(* IEC 61131-3 sources: plcassist-cli/packages/volt-lsp-iec/test-corpus/CodesysTestProject/Device/Plc Logic/Application/Library Manager/Standard, 22 files *)

(* ---- CONCAT.fun ---- *)
FUNCTION CONCAT : STRING(255)
VAR_INPUT
	STR1 : STRING(255);
	STR2 : STRING(255);
END_VAR
END_FUNCTION

(* ---- DELETE.fun ---- *)
FUNCTION DELETE : STRING(255)
VAR_INPUT
	STR : STRING(255);
	LEN : INT;
	POS : INT;
END_VAR
END_FUNCTION

(* ---- FIND.fun ---- *)
FUNCTION FIND : INT
VAR_INPUT
	STR1 : STRING(255);
	STR2 : STRING(255);
END_VAR
END_FUNCTION

(* ---- INSERT.fun ---- *)
FUNCTION INSERT : STRING(255)
VAR_INPUT
	STR1 : STRING(255);
	STR2 : STRING(255);
	POS : INT;
END_VAR
END_FUNCTION

(* ---- LEFT.fun ---- *)
FUNCTION LEFT : STRING(255)
VAR_INPUT
	STR : STRING(255);
	SIZE : INT;
END_VAR
END_FUNCTION

(* ---- LEN.fun ---- *)
FUNCTION LEN : INT
VAR_INPUT
	STR : STRING(255);
END_VAR
END_FUNCTION

(* ---- LEN_INTERNAL.fun ---- *)
FUNCTION LEN_INTERNAL : UINT
VAR_IN_OUT
	STR : STRING(255);
END_VAR
END_FUNCTION

(* ---- MEMCOPY_INTERNAL.fun ---- *)
FUNCTION MEMCOPY_INTERNAL : POINTER TO BYTE
VAR_INPUT
	PDEST : POINTER TO BYTE;
	PSRC : POINTER TO BYTE;
	DWSIZE : DWORD;
END_VAR
END_FUNCTION

(* ---- MID.fun ---- *)
FUNCTION MID : STRING(255)
VAR_INPUT
	STR : STRING(255);
	LEN : INT;
	POS : INT;
END_VAR
END_FUNCTION

(* ---- REPLACE.fun ---- *)
FUNCTION REPLACE : STRING(255)
VAR_INPUT
	STR1 : STRING(255);
	STR2 : STRING(255);
	L : INT;
	P : INT;
END_VAR
END_FUNCTION

(* ---- RIGHT.fun ---- *)
FUNCTION RIGHT : STRING(255)
VAR_INPUT
	STR : STRING(255);
	SIZE : INT;
END_VAR
END_FUNCTION

(* ---- CTD.fb ---- *)
FUNCTION_BLOCK CTD
VAR_INPUT
	CD : BOOL;
	LOAD : BOOL;
	PV : WORD;
END_VAR
VAR_OUTPUT
	Q : BOOL;
	CV : WORD;
END_VAR
VAR
	M : BOOL;
END_VAR
END_FUNCTION_BLOCK

(* ---- CTU.fb ---- *)
FUNCTION_BLOCK CTU
VAR_INPUT
	CU : BOOL;
	RESET : BOOL;
	PV : WORD;
END_VAR
VAR_OUTPUT
	Q : BOOL;
	CV : WORD;
END_VAR
VAR
	M : BOOL;
END_VAR
END_FUNCTION_BLOCK

(* ---- CTUD.fb ---- *)
FUNCTION_BLOCK CTUD
VAR_INPUT
	CU : BOOL;
	CD : BOOL;
	RESET : BOOL;
	LOAD : BOOL;
	PV : WORD;
END_VAR
VAR_OUTPUT
	QU : BOOL;
	QD : BOOL;
	CV : WORD;
END_VAR
VAR
	MU : BOOL;
	MD : BOOL;
	RU : BOOL;
	RD : BOOL;
END_VAR
END_FUNCTION_BLOCK

(* ---- F_TRIG.fb ---- *)
FUNCTION_BLOCK F_TRIG
VAR_INPUT
	CLK : BOOL;
END_VAR
VAR_OUTPUT
	Q : BOOL;
END_VAR
VAR
	M : BOOL := TRUE;
END_VAR
END_FUNCTION_BLOCK

(* ---- R_TRIG.fb ---- *)
FUNCTION_BLOCK R_TRIG
VAR_INPUT
	CLK : BOOL;
END_VAR
VAR_OUTPUT
	Q : BOOL;
END_VAR
VAR
	M : BOOL;
END_VAR
END_FUNCTION_BLOCK

(* ---- RS.fb ---- *)
FUNCTION_BLOCK RS
VAR_INPUT
	SET : BOOL;
	RESET1 : BOOL;
END_VAR
VAR_OUTPUT
	Q1 : BOOL;
END_VAR
END_FUNCTION_BLOCK

(* ---- RTC.fb ---- *)
FUNCTION_BLOCK RTC
VAR_INPUT
	EN : BOOL;
	PDT : DATE_AND_TIME;
END_VAR
VAR_OUTPUT
	Q : BOOL;
	CDT : DATE_AND_TIME;
END_VAR
VAR
	M : BOOL;
	DIFFTIME : TIME;
	LASTTIME : TIME := TIME#0ms;
	TIMEOFFSET : TIME := TIME#0ms;
	CURTIME : TIME;
END_VAR
END_FUNCTION_BLOCK

(* ---- SR.fb ---- *)
FUNCTION_BLOCK SR
VAR_INPUT
	SET1 : BOOL;
	RESET : BOOL;
END_VAR
VAR_OUTPUT
	Q1 : BOOL;
END_VAR
END_FUNCTION_BLOCK

(* ---- TOF.fb ---- *)
FUNCTION_BLOCK TOF
VAR_INPUT
	IN : BOOL;
	PT : TIME;
END_VAR
VAR_OUTPUT
	Q : BOOL;
	ET : TIME;
END_VAR
VAR
	M : BOOL;
	STARTTIME : TIME;
END_VAR
END_FUNCTION_BLOCK

(* ---- TON.fb ---- *)
FUNCTION_BLOCK TON
VAR_INPUT
	IN : BOOL;
	PT : TIME;
END_VAR
VAR_OUTPUT
	Q : BOOL;
	ET : TIME;
END_VAR
VAR
	M : BOOL;
	STARTTIME : TIME;
END_VAR
END_FUNCTION_BLOCK

(* ---- TP.fb ---- *)
FUNCTION_BLOCK TP
VAR_INPUT
	IN : BOOL;
	PT : TIME;
END_VAR
VAR_OUTPUT
	Q : BOOL;
	ET : TIME;
END_VAR
VAR
	STARTTIME : TIME;
END_VAR
END_FUNCTION_BLOCK
